{region 'Documentation'}
(*!
<summary>Checks inequality with the forbidden UINT value.</summary>
*)
{endregion}
FUNCTION_BLOCK AssertNotEqual_UInt EXTENDS AssertionBase
VAR_INPUT
    IN : UINT; //! Actual value checked or observed by this Assertion.
    Expected : UINT; //! Value that must differ from IN under this Assertion's comparison rules.
END_VAR

SUPER^();

{region 'Documentation'}
(*!
<summary>Check inequality with the forbidden UINT value.</summary>
*)
{endregion}
METHOD PROTECTED Assert
VAR
    Message : STRING(GVL_Constants.MessageLength);
    ExpectedText : STRING(GVL_Constants.AssertionValueLength);
    ActualText : STRING(GVL_Constants.AssertionValueLength);
END_VAR
IF NOT EvaluationActive THEN
    RETURN;
END_IF;

IF Result = E_Result.Error THEN
    RETURN;
END_IF;

IF Result = E_Result.Failed THEN
    RETURN;
END_IF;

IF IN = Expected THEN
    ExpectedText := UINT_TO_STRING(Expected);
    ActualText := UINT_TO_STRING(IN);
    Message := CONCAT('Assertion failed: values are equal but should differ. NotExpected = ',
        ExpectedText);
    Message := CONCAT(Message, ', Actual = ');
    Message := CONCAT(Message, ActualText);
    Message := CONCAT(Message, '.');
    Fail(Message := Message);
    RETURN;
END_IF;

Pass();
END_METHOD

END_FUNCTION_BLOCK

(* stored: Version 1.1.0.1
   POU AssertNotEqual_UInt: Id {6eadc651-b957-4f0a-b6ed-f213bae7102b}, SpecialFunc None
   Folder Internal: Id {f7460dfb-b001-4867-8c4a-2540e5d9c88a}
   Method Assert: Id {c4504d29-eec0-42e6-b6ce-6dbbcfdac7d0} *)
